// TwinCAT 3 PLC project ModeManagerCoreTests
// ProgramVersion: 3.1.4026.22
// libraries:
//   Tc2_Standard, * (Beckhoff Automation GmbH)
//   Tc2_System, * (Beckhoff Automation GmbH)
// project tree:
//   StateMachineControl/DUTs/ E_ModeState.TcDUT, ST_ModeManagerActions.TcDUT
//   StateMachineControl/POUs/ FB_HeartbeatWatchdog.TcPOU, FB_ModeManagerCore.TcPOU
//   StateMachineControl/tests/POUs/ PRG_ModeManagerCoreTests.TcPOU
//   StateMachineControl/tests/ ModeManagerCoreTestTask.TcTTO
// (motion and I/O tree: see PLC project experimentsequencertests)
// real-time tasks:
//   TASK DriveStateTestTask: cycle T#10ms, priority 1, ADS port 350
//   TASK TestTask: cycle T#10ms, priority 2, ADS port 351

CONFIGURATION ModeManagerCoreTests
    RESOURCE PLC ON TwinCAT3
        TASK ModeManagerCoreTestTask(INTERVAL := T#10ms, PRIORITY := 1);
        PROGRAM PRG_ModeManagerCoreTests WITH ModeManagerCoreTestTask : PRG_ModeManagerCoreTests;
    END_RESOURCE
END_CONFIGURATION

// ---- StateMachineControl/DUTs/E_ModeState.TcDUT
{attribute 'qualified_only'}
{attribute 'strict'}
{attribute 'to_string'}
TYPE E_ModeState :
(
    IDLE := 0,              // Servo OFF / initial
    RESETTING := 10,        // Reset pulse active — no experiment transitions allowed
    SERVO_READY := 20,      // Servo ON + drive OPERATION_ENABLED, awaiting experiment
    RUNNING := 30,          // Experiment active
    DONE := 40              // Playback complete, awaiting rearm
);
END_TYPE

// ---- StateMachineControl/DUTs/ST_ModeManagerActions.TcDUT
TYPE ST_ModeManagerActions :
STRUCT
    consumeResetReq : BOOL;
    clearModeFlags : BOOL;
    incrementResetAckCounter : BOOL;
    incrementWatchdogTripCounter : BOOL;
END_STRUCT
END_TYPE

// ---- StateMachineControl/tests/POUs/PRG_ModeManagerCoreTests.TcPOU
PROGRAM PRG_ModeManagerCoreTests
VAR
    lifecycleCore : FB_ModeManagerCore;
    doneCore : FB_ModeManagerCore;
    priorityCore : FB_ModeManagerCore;
    resetCore : FB_ModeManagerCore;
    staleStartCore : FB_ModeManagerCore;
    watchdogCore : FB_ModeManagerCore;
    simultaneousCore : FB_ModeManagerCore;
    testsExecuted : BOOL := FALSE;
    testsPassed : BOOL := FALSE;
    failureCount : UDINT := 0;
END_VAR

IF NOT testsExecuted THEN
    (* Cold IDLE and latched start waiting for both readiness inputs. *)
    lifecycleCore(servoEnableRequest := FALSE, experimentStartRequest := FALSE, anyModeRequest := FALSE, resetRequest := FALSE, experimentActivePreviousScan := FALSE, hostHeartbeatCounter := 0, heartbeatTimeoutTicks := 3, driveReadyPreviousScan := FALSE, loggerReady := FALSE, seqPlaybackDone := FALSE);
    IF (lifecycleCore.modeState <> E_ModeState.IDLE) OR lifecycleCore.driveEnable
        OR lifecycleCore.watchdogArmed OR lifecycleCore.watchdogTimeout THEN
        failureCount := failureCount + 1;
    END_IF

    lifecycleCore(servoEnableRequest := TRUE, experimentStartRequest := FALSE, anyModeRequest := TRUE, resetRequest := FALSE, experimentActivePreviousScan := FALSE, hostHeartbeatCounter := 1, heartbeatTimeoutTicks := 50, driveReadyPreviousScan := FALSE, loggerReady := FALSE, seqPlaybackDone := FALSE);
    IF (lifecycleCore.modeState <> E_ModeState.SERVO_READY) OR NOT lifecycleCore.driveEnable THEN
        failureCount := failureCount + 1;
    END_IF
    lifecycleCore(servoEnableRequest := TRUE, experimentStartRequest := TRUE, anyModeRequest := TRUE, resetRequest := FALSE, experimentActivePreviousScan := FALSE, hostHeartbeatCounter := 2, heartbeatTimeoutTicks := 50, driveReadyPreviousScan := FALSE, loggerReady := FALSE, seqPlaybackDone := FALSE);
    lifecycleCore(servoEnableRequest := TRUE, experimentStartRequest := FALSE, anyModeRequest := TRUE, resetRequest := FALSE, experimentActivePreviousScan := FALSE, hostHeartbeatCounter := 3, heartbeatTimeoutTicks := 50, driveReadyPreviousScan := TRUE, loggerReady := FALSE, seqPlaybackDone := FALSE);
    IF lifecycleCore.modeState <> E_ModeState.SERVO_READY THEN
        failureCount := failureCount + 1;
    END_IF
    lifecycleCore(servoEnableRequest := TRUE, experimentStartRequest := FALSE, anyModeRequest := TRUE, resetRequest := FALSE, experimentActivePreviousScan := FALSE, hostHeartbeatCounter := 4, heartbeatTimeoutTicks := 50, driveReadyPreviousScan := TRUE, loggerReady := TRUE, seqPlaybackDone := FALSE);
    IF (lifecycleCore.modeState <> E_ModeState.RUNNING) OR NOT lifecycleCore.driveEnable THEN
        failureCount := failureCount + 1;
    END_IF

    (* Explicit abort clears mode flags without a watchdog trip. *)
    lifecycleCore(servoEnableRequest := FALSE, experimentStartRequest := FALSE, anyModeRequest := FALSE, resetRequest := FALSE, experimentActivePreviousScan := TRUE, hostHeartbeatCounter := 5, heartbeatTimeoutTicks := 50, driveReadyPreviousScan := TRUE, loggerReady := TRUE, seqPlaybackDone := FALSE);
    IF (lifecycleCore.modeState <> E_ModeState.IDLE) OR lifecycleCore.driveEnable
        OR NOT lifecycleCore.actions.clearModeFlags
        OR lifecycleCore.actions.incrementWatchdogTripCounter THEN
        failureCount := failureCount + 1;
    END_IF
    lifecycleCore(servoEnableRequest := FALSE, experimentStartRequest := FALSE, anyModeRequest := FALSE, resetRequest := FALSE, experimentActivePreviousScan := FALSE, hostHeartbeatCounter := 6, heartbeatTimeoutTicks := 50, driveReadyPreviousScan := TRUE, loggerReady := TRUE, seqPlaybackDone := FALSE);
    IF lifecycleCore.actions.clearModeFlags THEN
        failureCount := failureCount + 1;
    END_IF

    (* Natural completion latches DONE until an explicit reset, so ADS polling cannot miss it. *)
    doneCore(servoEnableRequest := TRUE, experimentStartRequest := FALSE, anyModeRequest := TRUE, resetRequest := FALSE, experimentActivePreviousScan := FALSE, hostHeartbeatCounter := 1, heartbeatTimeoutTicks := 50, driveReadyPreviousScan := FALSE, loggerReady := FALSE, seqPlaybackDone := FALSE);
    doneCore(servoEnableRequest := TRUE, experimentStartRequest := TRUE, anyModeRequest := TRUE, resetRequest := FALSE, experimentActivePreviousScan := FALSE, hostHeartbeatCounter := 2, heartbeatTimeoutTicks := 50, driveReadyPreviousScan := TRUE, loggerReady := TRUE, seqPlaybackDone := FALSE);
    doneCore(servoEnableRequest := TRUE, experimentStartRequest := FALSE, anyModeRequest := TRUE, resetRequest := FALSE, experimentActivePreviousScan := TRUE, hostHeartbeatCounter := 3, heartbeatTimeoutTicks := 50, driveReadyPreviousScan := TRUE, loggerReady := TRUE, seqPlaybackDone := TRUE);
    IF (doneCore.modeState <> E_ModeState.DONE) OR doneCore.driveEnable
        OR NOT doneCore.actions.clearModeFlags THEN
        failureCount := failureCount + 1;
    END_IF
    doneCore(servoEnableRequest := FALSE, experimentStartRequest := FALSE, anyModeRequest := FALSE, resetRequest := FALSE, experimentActivePreviousScan := FALSE, hostHeartbeatCounter := 4, heartbeatTimeoutTicks := 50, driveReadyPreviousScan := TRUE, loggerReady := TRUE, seqPlaybackDone := FALSE);
    IF doneCore.modeState <> E_ModeState.DONE THEN
        failureCount := failureCount + 1;
    END_IF
    doneCore(servoEnableRequest := FALSE, experimentStartRequest := FALSE, anyModeRequest := FALSE, resetRequest := TRUE, experimentActivePreviousScan := FALSE, hostHeartbeatCounter := 5, heartbeatTimeoutTicks := 50, driveReadyPreviousScan := TRUE, loggerReady := TRUE, seqPlaybackDone := FALSE);
    IF doneCore.modeState <> E_ModeState.RESETTING THEN
        failureCount := failureCount + 1;
    END_IF

    (* Drive loss wins over simultaneous sequence completion. *)
    priorityCore(servoEnableRequest := TRUE, experimentStartRequest := FALSE, anyModeRequest := TRUE, resetRequest := FALSE, experimentActivePreviousScan := FALSE, hostHeartbeatCounter := 1, heartbeatTimeoutTicks := 50, driveReadyPreviousScan := FALSE, loggerReady := FALSE, seqPlaybackDone := FALSE);
    priorityCore(servoEnableRequest := TRUE, experimentStartRequest := TRUE, anyModeRequest := TRUE, resetRequest := FALSE, experimentActivePreviousScan := FALSE, hostHeartbeatCounter := 2, heartbeatTimeoutTicks := 50, driveReadyPreviousScan := TRUE, loggerReady := TRUE, seqPlaybackDone := FALSE);
    priorityCore(servoEnableRequest := TRUE, experimentStartRequest := FALSE, anyModeRequest := TRUE, resetRequest := FALSE, experimentActivePreviousScan := TRUE, hostHeartbeatCounter := 3, heartbeatTimeoutTicks := 50, driveReadyPreviousScan := FALSE, loggerReady := TRUE, seqPlaybackDone := TRUE);
    IF (priorityCore.modeState <> E_ModeState.IDLE) OR NOT priorityCore.actions.clearModeFlags THEN
        failureCount := failureCount + 1;
    END_IF

    (* hold=1 means RESETTING on the edge call and one additional call. *)
    resetCore(servoEnableRequest := TRUE, experimentStartRequest := TRUE, anyModeRequest := TRUE, resetRequest := TRUE, experimentActivePreviousScan := FALSE, hostHeartbeatCounter := 1, heartbeatTimeoutTicks := 50, driveReadyPreviousScan := TRUE, loggerReady := TRUE, seqPlaybackDone := FALSE);
    IF (resetCore.modeState <> E_ModeState.RESETTING)
        OR NOT resetCore.actions.consumeResetReq
        OR NOT resetCore.actions.clearModeFlags
        OR NOT resetCore.actions.incrementResetAckCounter
        OR resetCore.actions.incrementWatchdogTripCounter THEN
        failureCount := failureCount + 1;
    END_IF
    resetCore(servoEnableRequest := FALSE, experimentStartRequest := FALSE, anyModeRequest := FALSE, resetRequest := TRUE, experimentActivePreviousScan := FALSE, hostHeartbeatCounter := 2, heartbeatTimeoutTicks := 50, driveReadyPreviousScan := TRUE, loggerReady := TRUE, seqPlaybackDone := FALSE);
    IF (resetCore.modeState <> E_ModeState.RESETTING)
        OR resetCore.actions.consumeResetReq OR resetCore.actions.incrementResetAckCounter THEN
        failureCount := failureCount + 1;
    END_IF
    resetCore(servoEnableRequest := FALSE, experimentStartRequest := FALSE, anyModeRequest := FALSE, resetRequest := TRUE, experimentActivePreviousScan := FALSE, hostHeartbeatCounter := 3, heartbeatTimeoutTicks := 50, driveReadyPreviousScan := TRUE, loggerReady := TRUE, seqPlaybackDone := FALSE);
    IF (resetCore.modeState <> E_ModeState.IDLE)
        OR resetCore.actions.consumeResetReq OR resetCore.actions.incrementResetAckCounter THEN
        failureCount := failureCount + 1;
    END_IF
    resetCore(servoEnableRequest := FALSE, experimentStartRequest := FALSE, anyModeRequest := FALSE, resetRequest := FALSE, experimentActivePreviousScan := FALSE, hostHeartbeatCounter := 4, heartbeatTimeoutTicks := 50, driveReadyPreviousScan := TRUE, loggerReady := TRUE, seqPlaybackDone := FALSE);
    resetCore(servoEnableRequest := FALSE, experimentStartRequest := FALSE, anyModeRequest := FALSE, resetRequest := TRUE, experimentActivePreviousScan := FALSE, hostHeartbeatCounter := 5, heartbeatTimeoutTicks := 50, driveReadyPreviousScan := TRUE, loggerReady := TRUE, seqPlaybackDone := FALSE);
    IF NOT resetCore.actions.consumeResetReq OR NOT resetCore.actions.incrementResetAckCounter THEN
        failureCount := failureCount + 1;
    END_IF

    (* A start edge observed during RESETTING must not survive an explicit abort. *)
    staleStartCore(servoEnableRequest := FALSE, experimentStartRequest := FALSE, anyModeRequest := FALSE, resetRequest := TRUE, experimentActivePreviousScan := FALSE, hostHeartbeatCounter := 1, heartbeatTimeoutTicks := 50, driveReadyPreviousScan := FALSE, loggerReady := FALSE, seqPlaybackDone := FALSE);
    staleStartCore(servoEnableRequest := TRUE, experimentStartRequest := TRUE, anyModeRequest := TRUE, resetRequest := FALSE, experimentActivePreviousScan := FALSE, hostHeartbeatCounter := 2, heartbeatTimeoutTicks := 50, driveReadyPreviousScan := TRUE, loggerReady := TRUE, seqPlaybackDone := FALSE);
    staleStartCore(servoEnableRequest := FALSE, experimentStartRequest := FALSE, anyModeRequest := FALSE, resetRequest := FALSE, experimentActivePreviousScan := FALSE, hostHeartbeatCounter := 3, heartbeatTimeoutTicks := 50, driveReadyPreviousScan := TRUE, loggerReady := TRUE, seqPlaybackDone := FALSE);
    IF staleStartCore.modeState <> E_ModeState.IDLE THEN
        failureCount := failureCount + 1;
    END_IF
    staleStartCore(servoEnableRequest := TRUE, experimentStartRequest := FALSE, anyModeRequest := TRUE, resetRequest := FALSE, experimentActivePreviousScan := FALSE, hostHeartbeatCounter := 4, heartbeatTimeoutTicks := 50, driveReadyPreviousScan := TRUE, loggerReady := TRUE, seqPlaybackDone := FALSE);
    staleStartCore(servoEnableRequest := TRUE, experimentStartRequest := FALSE, anyModeRequest := TRUE, resetRequest := FALSE, experimentActivePreviousScan := FALSE, hostHeartbeatCounter := 5, heartbeatTimeoutTicks := 50, driveReadyPreviousScan := TRUE, loggerReady := TRUE, seqPlaybackDone := FALSE);
    IF (staleStartCore.modeState <> E_ModeState.SERVO_READY) OR NOT staleStartCore.driveEnable THEN
        failureCount := failureCount + 1;
    END_IF

    (* Timeout occurs on the configured armed call and trips only once. *)
    watchdogCore(servoEnableRequest := FALSE, experimentStartRequest := FALSE, anyModeRequest := FALSE, resetRequest := FALSE, experimentActivePreviousScan := FALSE, hostHeartbeatCounter := 10, heartbeatTimeoutTicks := 2, driveReadyPreviousScan := FALSE, loggerReady := FALSE, seqPlaybackDone := FALSE);
    watchdogCore(servoEnableRequest := TRUE, experimentStartRequest := FALSE, anyModeRequest := TRUE, resetRequest := FALSE, experimentActivePreviousScan := FALSE, hostHeartbeatCounter := 10, heartbeatTimeoutTicks := 2, driveReadyPreviousScan := FALSE, loggerReady := FALSE, seqPlaybackDone := FALSE);
    IF watchdogCore.watchdogTimeout OR (watchdogCore.modeState <> E_ModeState.SERVO_READY) THEN
        failureCount := failureCount + 1;
    END_IF
    watchdogCore(servoEnableRequest := TRUE, experimentStartRequest := FALSE, anyModeRequest := TRUE, resetRequest := FALSE, experimentActivePreviousScan := FALSE, hostHeartbeatCounter := 10, heartbeatTimeoutTicks := 2, driveReadyPreviousScan := FALSE, loggerReady := FALSE, seqPlaybackDone := FALSE);
    IF NOT watchdogCore.watchdogTimeout OR NOT watchdogCore.actions.incrementWatchdogTripCounter
        OR NOT watchdogCore.actions.clearModeFlags OR (watchdogCore.modeState <> E_ModeState.IDLE) THEN
        failureCount := failureCount + 1;
    END_IF
    watchdogCore(servoEnableRequest := TRUE, experimentStartRequest := FALSE, anyModeRequest := TRUE, resetRequest := FALSE, experimentActivePreviousScan := FALSE, hostHeartbeatCounter := 10, heartbeatTimeoutTicks := 2, driveReadyPreviousScan := FALSE, loggerReady := FALSE, seqPlaybackDone := FALSE);
    IF NOT watchdogCore.watchdogTimeout OR watchdogCore.actions.incrementWatchdogTripCounter THEN
        failureCount := failureCount + 1;
    END_IF

    (* Watchdog wins over reset, but the reset request is still consumed. *)
    simultaneousCore(servoEnableRequest := TRUE, experimentStartRequest := FALSE, anyModeRequest := TRUE, resetRequest := TRUE, experimentActivePreviousScan := FALSE, hostHeartbeatCounter := 0, heartbeatTimeoutTicks := 0, driveReadyPreviousScan := FALSE, loggerReady := FALSE, seqPlaybackDone := FALSE);
    IF (simultaneousCore.modeState <> E_ModeState.IDLE)
        OR NOT simultaneousCore.actions.consumeResetReq
        OR NOT simultaneousCore.actions.clearModeFlags
        OR simultaneousCore.actions.incrementResetAckCounter
        OR NOT simultaneousCore.actions.incrementWatchdogTripCounter THEN
        failureCount := failureCount + 1;
    END_IF

    testsExecuted := TRUE;
    testsPassed := (failureCount = 0);
END_IF

END_PROGRAM

// ---- StateMachineControl/POUs/FB_ModeManagerCore.TcPOU
FUNCTION_BLOCK FB_ModeManagerCore
VAR_INPUT
    servoEnableRequest : BOOL;
    experimentStartRequest : BOOL;
    anyModeRequest : BOOL;
    resetRequest : BOOL;
    experimentActivePreviousScan : BOOL;
    hostHeartbeatCounter : UDINT;
    heartbeatTimeoutTicks : UDINT;
    driveReadyPreviousScan : BOOL;
    loggerReady : BOOL;
    seqPlaybackDone : BOOL;
END_VAR
VAR_OUTPUT
    modeState : E_ModeState := E_ModeState.IDLE;
    driveEnable : BOOL := FALSE;
    watchdogArmed : BOOL := FALSE;
    watchdogTimeout : BOOL := FALSE;
    actions : ST_ModeManagerActions;
END_VAR
VAR
    servoEnableRequestPrev : BOOL := FALSE;
    experimentStartRequestPrev : BOOL := FALSE;
    servoEnableEdge : BOOL := FALSE;
    experimentStartEdge : BOOL := FALSE;
    servoEnableLatched : BOOL := FALSE;
    experimentStartLatched : BOOL := FALSE;
    resetRequestPrev : BOOL := FALSE;
    resetEdge : BOOL := FALSE;
    resetHoldTicksRemaining : UDINT := 0;
    fbHeartbeatWatchdog : FB_HeartbeatWatchdog;
END_VAR
VAR CONSTANT
    RESET_PULSE_HOLD_TICKS : UDINT := 1;
END_VAR

actions.consumeResetReq := FALSE;
actions.clearModeFlags := FALSE;
actions.incrementResetAckCounter := FALSE;
actions.incrementWatchdogTripCounter := FALSE;

servoEnableEdge := servoEnableRequest AND NOT servoEnableRequestPrev;
experimentStartEdge := experimentStartRequest AND NOT experimentStartRequestPrev;
servoEnableRequestPrev := servoEnableRequest;
experimentStartRequestPrev := experimentStartRequest;

IF servoEnableEdge THEN
    servoEnableLatched := TRUE;
END_IF
IF experimentStartEdge THEN
    experimentStartLatched := TRUE;
END_IF
(* A missing servo request is the explicit abort contract.  Clear both
   latches so a start captured during RESETTING cannot run after rearm. *)
IF NOT servoEnableRequest THEN
    servoEnableLatched := FALSE;
    experimentStartLatched := FALSE;
END_IF

resetEdge := resetRequest AND NOT resetRequestPrev;
IF resetEdge THEN
    actions.consumeResetReq := TRUE;
END_IF
resetRequestPrev := resetRequest;

watchdogArmed := anyModeRequest OR experimentActivePreviousScan OR servoEnableLatched;
fbHeartbeatWatchdog(
    enable := watchdogArmed,
    heartbeatCounter := hostHeartbeatCounter,
    timeoutTicks := heartbeatTimeoutTicks
);
watchdogTimeout := fbHeartbeatWatchdog.timeout;

IF watchdogTimeout THEN
    modeState := E_ModeState.IDLE;
    actions.clearModeFlags := TRUE;
    servoEnableLatched := FALSE;
    experimentStartLatched := FALSE;
    IF fbHeartbeatWatchdog.tripEdge THEN
        actions.incrementWatchdogTripCounter := TRUE;
    END_IF

ELSIF resetEdge THEN
    modeState := E_ModeState.RESETTING;
    resetHoldTicksRemaining := RESET_PULSE_HOLD_TICKS;
    actions.clearModeFlags := TRUE;
    actions.incrementResetAckCounter := TRUE;
    servoEnableLatched := FALSE;
    experimentStartLatched := FALSE;

ELSE
    CASE modeState OF
        E_ModeState.IDLE:
            IF servoEnableLatched THEN
                modeState := E_ModeState.SERVO_READY;
            END_IF

        E_ModeState.RESETTING:
            IF resetHoldTicksRemaining > 0 THEN
                resetHoldTicksRemaining := resetHoldTicksRemaining - 1;
            ELSE
                modeState := E_ModeState.IDLE;
            END_IF

        E_ModeState.SERVO_READY:
            IF NOT servoEnableLatched THEN
                modeState := E_ModeState.IDLE;
                experimentStartLatched := FALSE;
            ELSIF experimentStartLatched AND driveReadyPreviousScan AND loggerReady THEN
                modeState := E_ModeState.RUNNING;
                experimentStartLatched := FALSE;
            END_IF

        E_ModeState.RUNNING:
            IF NOT servoEnableLatched OR NOT driveReadyPreviousScan THEN
                modeState := E_ModeState.IDLE;
                experimentStartLatched := FALSE;
                servoEnableLatched := FALSE;
                actions.clearModeFlags := TRUE;
            ELSIF seqPlaybackDone THEN
                modeState := E_ModeState.DONE;
                servoEnableLatched := FALSE;
                experimentStartLatched := FALSE;
                actions.clearModeFlags := TRUE;
            END_IF

        E_ModeState.DONE:
            servoEnableLatched := FALSE;
            experimentStartLatched := FALSE;
    END_CASE
END_IF

driveEnable := servoEnableLatched
    AND (modeState = E_ModeState.SERVO_READY OR modeState = E_ModeState.RUNNING);

END_FUNCTION_BLOCK

// ---- StateMachineControl/POUs/FB_HeartbeatWatchdog.TcPOU
FUNCTION_BLOCK FB_HeartbeatWatchdog
VAR_INPUT
    enable : BOOL;
    heartbeatCounter : UDINT;
    timeoutTicks : UDINT;
END_VAR
VAR_OUTPUT
    timeout : BOOL := FALSE;
    tripEdge : BOOL := FALSE;
END_VAR
VAR
    counterPrev : UDINT := 0;
    silenceTicks : UDINT := 0;
    tripLatched : BOOL := FALSE;
    heartbeatChanged : BOOL := FALSE;
END_VAR

tripEdge := FALSE;
heartbeatChanged := (heartbeatCounter <> counterPrev);

IF NOT enable THEN
    counterPrev := heartbeatCounter;
    silenceTicks := 0;
    tripLatched := FALSE;
ELSIF heartbeatChanged THEN
    counterPrev := heartbeatCounter;
    silenceTicks := 0;
    tripLatched := FALSE;
ELSE
    IF silenceTicks < timeoutTicks THEN
        silenceTicks := silenceTicks + 1;
    END_IF
END_IF

timeout := enable AND (silenceTicks >= timeoutTicks);
IF timeout AND NOT tripLatched THEN
    tripEdge := TRUE;
    tripLatched := TRUE;
END_IF

END_FUNCTION_BLOCK
